Staubli VAL3: _onStartPROG.pgx

public program _onStartPROG(string x_sHtml)
begin
  nPgIndexPROG=0
  nPgNumPROG=0
  sPagePROG=""
  sPgIndexPROG=""
  bSelProg=true
  bSelTraj=false
  if bSelProg
    call resfreshPROG(x_sHtml)
  elseIf bSelTraj
    call resfreshTRAJ(x_sHtml)
  endIf
end
